           REGION Request selector
               //set Index and RecordLen based on the request
               IF #statParameterPage0 THEN
                   #statIndex := #INDEX_DIRECT_PARAM0;
                   #statRecordLen := #LENGTH_DIRECT_PARAM0;
               ELSIF #statSystemCommands THEN
                   #statIndex := #INDEX_SYSTEM_COMMANDS;
                   #statRecordLen := #LENGTH_SYSTEM_COMMANDS;
               ELSIF #statVendorName THEN
                   #statIndex := #INDEX_VENDOR_NAME;
                   #statRecordLen := #LENGTH_VENDOR_NAME;
               ELSIF #statVendorText THEN
                   #statIndex := #INDEX_VENDOR_TEXT;
                   #statRecordLen := #LENGTH_VENDOR_TEXT;
               ELSIF #statProductName THEN
                   #statIndex := #INDEX_PRODUCT_NAME;
                   #statRecordLen := #LENGTH_PRODUCT_NAME;
               ELSIF #statProductID THEN
                   #statIndex := #INDEX_PRODUCT_ID;
                   #statRecordLen := #LENGTH_PRODUCT_ID;
               ELSIF #statHwRevision THEN
                   #statIndex := #INDEX_HARDWARE_REVISION;
                   #statRecordLen := #LENGTH_HARDWARE_REVISION;
               ELSIF #statFwRevision THEN
                   #statIndex := #INDEX_FIRMWARE_REVISION;
                   #statRecordLen := #LENGTH_FIRMWARE_REVISION;
               ELSIF #statAppSpecificName THEN
                   #statIndex := #INDEX_APP_SPECIFIC_NAME;
                   #statRecordLen := #LENGTH_APP_SPECIFIC_NAME;
               ELSIF #statDiagnosis THEN
                   #statIndex := #INDEX_DIAGNOSTICS;
                   #statRecordLen := #LENGTH_DIAGNOSTICS;
               ELSIF #statMeasurements THEN
                   #statIndex := #INDEX_MEASUREMENTS;
                   #statRecordLen := #LENGTH_MEASUREMENTS;
               ELSIF #statParameters THEN
                   #statIndex := #INDEX_PARAMETERS;
                   #statRecordLen := #LENGTH_PARAMETERS;
               ELSE
                   RETURN;
               END_IF;
           END_REGION

           IF #statReadWrite = #MODE_WRITE THEN
               //prepare statRecord in case of a writing request
               REGION write
                   IF #statSystemCommands THEN
                       #statRecord[0] := #data.systemCommands;

                   ELSIF #statAppSpecificName THEN
                       Strg_TO_Chars(Strg := #data.appSpecificName,
                                     pChars := 0,
                                     Cnt => #tempLen,
                                     Chars := #statRecord);

                       // Fill remaining characters with null
                       FOR #tempIndex := UINT_TO_INT(#tempLen) TO #statRecordLen - 1 DO
                           #statRecord[#tempIndex] := CHAR_TO_BYTE(#EMPTY_CHAR);
                       END_FOR;

                   ELSIF #statParameters THEN
                       #tempRetValSerialize := Serialize(SRC_VARIABLE := #data.parameters, DEST_ARRAY => #tempFieldParameters, POS := #tempPosSerialize);
                       UMOVE_BLK(IN := #tempFieldParameters[0],
                                 COUNT := INT_TO_ULINT(#statRecordLen),
                                 OUT => #statRecord[0]);
                   ELSE    // all other data set are read only
                       ;
                   END_IF;
                   #tempInternalError := #tempRetValSerialize <> WORD_TO_INT(#STATUS_EXECUTION_FINISHED);
               END_REGION

           END_IF;
       END_IF;
   END_REGION

   REGION CALL
       //IOL-Call -> Request to read/write from an IO-Link-Device
       #instDevice(execute := #execute,
                   hwID := #statHwID,
                   cap := #statCap,
                   readWrite := #statReadWrite,
                   "port" := #statPort,
                   pollingPeriod := #statPollingPeriod,
                   index := #statIndex,
                   subindex := #statSubindex,
                   writeLen := #statRecordLen,
                   timeout := #DEVICE_TIMEOUT,
                   record := #statRecord);
   END_REGION

   REGION READ
       // Copy data if available and valid
       IF #instDevice.done = TRUE AND #statDoneOld = FALSE AND #statReadWrite = #MODE_READ THEN
           IF #statParameterPage0 THEN
               UMOVE_BLK(IN := #statRecord[0],
                         COUNT := INT_TO_ULINT(#statRecordLen),
                         OUT => #tempFieldParameterPage0[0]);
               #tempRetValDeserialize := Deserialize(SRC_ARRAY := #tempFieldParameterPage0, DEST_VARIABLE => #data.parameterPage0, POS := #tempPosDeserialize);
           ELSIF #statVendorName THEN
               Chars_TO_Strg(Chars := #statRecord,
                             pChars := 0,
                             Cnt := INT_TO_UINT(#statRecordLen),
                             Strg => #data.vendorName);
           ELSIF #statVendorText THEN
               Chars_TO_Strg(Chars := #statRecord,
                             pChars := 0,
                             Cnt := INT_TO_UINT(#statRecordLen),
                             Strg => #data.vendorText);
           ELSIF #statProductName THEN
               Chars_TO_Strg(Chars := #statRecord,
                             pChars := 0,
                             Cnt := INT_TO_UINT(#statRecordLen),
                             Strg => #data.productName);
           ELSIF #statProductID THEN
               Chars_TO_Strg(Chars := #statRecord,
                             pChars := 0,
                             Cnt := INT_TO_UINT(#statRecordLen),
                             Strg => #data.productID);
           ELSIF #statHwRevision THEN
               Chars_TO_Strg(Chars := #statRecord,
                             pChars := 0,
                             Cnt := INT_TO_UINT(#statRecordLen),
                             Strg => #data.hwRevision);
           ELSIF #statFwRevision THEN
               Chars_TO_Strg(Chars := #statRecord,
                             pChars := 0,
                             Cnt := INT_TO_UINT(#statRecordLen),
                             Strg => #data.fwRevision);
           ELSIF #statAppSpecificName THEN
               Chars_TO_Strg(Chars := #statRecord,
                             pChars := 0,
                             Cnt := INT_TO_UINT(#statRecordLen),
                             Strg => #data.appSpecificName);
           ELSIF #statDiagnosis THEN
               UMOVE_BLK(IN := #statRecord[0],
                         COUNT := INT_TO_ULINT(#statRecordLen),
                         OUT => #tempFieldDiagnostics[0]);
               #tempRetValDeserialize := Deserialize(SRC_ARRAY := #tempFieldDiagnostics, DEST_VARIABLE => #data.diagnostics, POS := #tempPosDeserialize);
           ELSIF #statMeasurements THEN
               UMOVE_BLK(IN := #statRecord[0],
                         COUNT := INT_TO_ULINT(#statRecordLen),
                         OUT => #tempFieldMeasurements[0]);
               #tempRetValDeserialize := Deserialize(SRC_ARRAY := #tempFieldMeasurements, DEST_VARIABLE => #data.measuredValues, POS := #tempPosDeserialize);
           ELSIF #statParameters THEN
               UMOVE_BLK(IN := #statRecord[0],
                         COUNT := INT_TO_ULINT(#statRecordLen),
                         OUT => #tempFieldParameters[0]);
               #tempRetValDeserialize := Deserialize(SRC_ARRAY := #tempFieldParameters, DEST_VARIABLE => #data.parameters, POS := #tempPosDeserialize);
           ELSE  // Other data sets are not defined
               ;
           END_IF;
           #tempInternalError := #tempRetValDeserialize <> WORD_TO_INT(#STATUS_EXECUTION_FINISHED);
       END_IF;

       #statDoneOld := #instDevice.done;
   END_REGION

   REGION OUTPUTS
       IF #tempInternalError THEN //Error occured
           #done := false;
           #busy := false;
           #error := true;
           #status := #ERR_INCONSISTENT_DATA;
       ELSE //Execute successful
           #done := #instDevice.done;
           #busy := #instDevice.busy;
           #error := #instDevice.error;
           #status := #instDevice.status;
           #diagnostics := #instDevice.diagnostics;
       END_IF;
   END_REGION
END_FUNCTION_BLOCK

// folder: LIOLink/S7-1200/1500/Device-specific blocks/SIRIUS/SIRIUS WD

FUNCTION_BLOCK "LIOLink_8WD46"   // FB2, SCL
TITLE = LIOLink_8WD46
{ S7_Optimized_Access := 'TRUE' }
FAMILY : LIOLink
VERSION : 1.0
// Capsule block to communicate with 8WD46
   VAR_INPUT
      execute : Bool;   // Request to execute function
      hwID : HW_IO;   // Hardware identifier of IO-Link master module or first sub module
      cap : Int;   // Client Access Point (CAP) 0xB400 or 0x00E3 (227)
      readWrite : Bool;   // FALSE: read, TRUE: write
      port : Int;   // Port of the IO-Link Master for the Device
      pollingPeriod : Time := T#100MS;   // Time period of polling
      systemCommands : Bool;   // Write system commands
      vendorName : Bool;   // Read Vendor Name
      vendorText : Bool;   // Read Vendor Text
      productName : Bool;   // Read Product Name
      productID : Bool;   // Read Product ID
      productText : Bool;   // Read Product Text
      hwRevision : Bool;   // Read Hardware revision
      fwRevision : Bool;   // Read firmware revision
      appSpecificName : Bool;   // Read/Write Application Specific Name
      functionTag : Bool;   // Read/Write: function tag
      locationTag : Bool;   // Read/Write: location tag
      opHour : Bool;   // Read operating hour
      operatingMode : Bool;   // Read/Write: operating mode (signal mode, auto scale mode, ...)
      lightEffect : USInt;   // Read/Write light effect - 1 to 15: select segment
      soundMode : USInt;   // Read ID of the inserted ID key
      powerReduction : Bool;   // Read/Write power reduction (0: on / 1: off)
      fillLevelMode : Bool;   // Read/Write only in level mode (0: use settings of segment 1-9,15 / 1: use settings of segment 1 )
      headlong : Bool;   // Read/Write orientation of installation (normal / overhead)
      elementCount : Bool;   // Read/Write number of elements
   END_VAR
   VAR_OUTPUT
      done : Bool;   // TRUE: Commanded functionality has been completed successfully
      busy : Bool;   // TRUE: FB is not finished and new output values can be expected
      error : Bool;   // TRUE: An error occurred during the execution of the FB
      status : Word;   // 16#0000 - 16#7FFF: Status of the FB, 16#8000 - 16#FFFF: Error identification
      diagnostics : "LIOLink_typeDiagnostics";   // Diagnostics information of LIOLink_Device
   END_VAR
   VAR_IN_OUT
      data : "LIOLink_8WD46_typeAll";   // Data area, device specific (Data Type)
   END_VAR
   VAR
      instDevice : "LIOLink_Device";
      statRecord : Array[0..#UPPER_BOUND_RECORD] of Byte;   // Record buffer
      statIndex : Int;   // Requested index
      statSubindex : Int;   // Requested subindex
      statRecordLen : Int;   // Length of record to be written
      statHwID : HW_IO;   // Static value for input 'hwID'
      statCap : Int;   // Static value for input 'cap'
      statReadWrite : Bool;   // Static value for input 'readWrite'
      statPort : Int;   // Static value for input 'port'
      statPollingPeriod : Time;   // Static value for input 'pollingPeriod'
      statSystemCommands : Bool;   // Static value for input 'systemCommands'
      statVendorName : Bool;   // Static value for input 'vendorName'
      statVendorText : Bool;   // Static value for input 'vendorText'
      statProductName : Bool;   // Static value for input 'productName'
      statProductID : Bool;   // Static value for input 'productID'
      statProductText : Bool;   // Static value for input 'productText'
      statHwRevision : Bool;   // Static value for input 'hwRevision'
      statFwRevision : Bool;   // Static value for input 'fwRevision'
      statAppSpecificName : Bool;   // Static value for input 'appSpecificName'
      statFunctionTag : Bool;   // Static value for input 'functionTag'
      statLocationTag : Bool;   // Static value for input 'locationTag'
      statOpHour : Bool;   // Static value for input 'opHour'
      statOperatingMode : Bool;   // Static value for input 'operatingMode'
      statLightEffect : USInt;   // Static value for input 'lightEffect'
      statSoundMode : USInt;   // Static value for input 'soundMode'
      statPowerReduction : Bool;   // Static value for input 'powerReduction'
      statFillLevelMode : Bool;   // Static value for input 'fillLevelMode'
      statHeadlong : Bool;   // Static value for input 'headLong'
      statElementCount : Bool;   // Static value for input 'elementCount'
      statRequest : Int;   // Case of request (data set)
      statDoneOld : Bool;   // Last cycle's value of instDevice.done
   END_VAR
   VAR_TEMP
      tempIndex : Int;   // Loop index
      tempLen : UInt;   // Length
      tempRetValSerialize : Int;   // Auxiliary tag for Serialize RetVal
      tempRetValDeserialize : Int;   // Auxiliary tag for Deserialize RetVal
      tempPosSerialize : DInt;   // Auxiliary tag for Serialize POS Output
      tempPosDeserialize : DInt;   // Auxiliary tag for Deserialize POS Output
      tempFieldLightEffects : Array[0..#UPPER_BOUND_LIGHT_EFFECTS] of Byte;   // Auxiliary tag for Light Effects record conversion
      tempFieldSoundMode : Array[0..#UPPER_BOUND_SOUND_MODE] of Byte;   // Auxiliary tag for Sound Mode record conversion
      tempFieldOpHour : Array[0..#UPPER_BOUND_OP_HOUR] of Byte;   // Auxiliary tag for Op Hour record conversion
      tempFieldDiagnostics : Array[0..#UPPER_BOUND_DIAGNOSTICS] of Byte;   // Auxiliary tag for Diagnostics record conversion
      tempInternalError : Bool;   // Auxiliary tag to collect serialize and Deserialize issues
   END_VAR
   VAR CONSTANT
      UPPER_BOUND_RECORD : Int := 231;   // Upper Bound of record buffer
      HIGHEST_REQUEST_NUMBER : Int := 28;   // Highest available request number
      UPPER_BOUND_LIGHT_EFFECTS : Int := 7;   // Upper Bound of Light Effects auxiliary field
      UPPER_BOUND_SOUND_MODE : Int := 15;   // Upper Bound of Sound Mode auxiliary field
      UPPER_BOUND_OP_HOUR : Int := 3;   // Upper Bound of Op Hours auxiliary field
      UPPER_BOUND_DIAGNOSTICS : Int := 19;   // Upper Bound of Diagnostics auxiliary field
      MODE_READ : Bool := FALSE;   // Mode to read data
      MODE_WRITE : Bool := TRUE;   // Mode to write data
      STATUS_IDLE : Word := 16#7000;   // Status: Idle
      STATUS_EXECUTION_FINISHED : Word := 16#0000;   // Execution finished without errors
      ERR_INCONSISTENT_DATA : Word := 16#8402;   // Error: Read data record doesn't match request
      INDEX_SYSTEM_COMMANDS : Int := 2;   // Record Index
      INDEX_VENDOR_NAME : Int := 16;   // Record Index
      INDEX_VENDOR_TEXT : Int := 17;   // Record Index
      INDEX_PRODUCT_NAME : Int := 18;   // Record Index
      INDEX_PRODUCT_ID : Int := 19;   // Record Index
      INDEX_PRODUCT_TEXT : Int := 20;   // Record Index
      INDEX_HARDWARE_REVISION : Int := 22;   // Record Index
      INDEX_FIRMWARE_REVISION : Int := 23;   // Record Index
      INDEX_APP_SPECIFIC_NAME : Int := 24;   // Record Index
      INDEX_FUNCTION_TAG : Int := 25;   // Record Index
      INDEX_LOCATION_TAG : Int := 26;   // Record Index
      INDEX_OPERATING_HOURS : Int := 74;   // Record Index
      INDEX_OPERATING_MODE : Int := 100;   // Record Index
      INDEX_LIGHT_EFFECT : Int := 101;   // Record Index - start of range
      SEGMENT_COUNT_MAX : Int := 15;   // maximum count of segments
      INDEX_SOUND_MODE : Int := 120;   // Record Index - start of range
      SOUND_COUNT_MAX : Int := 10;   // maximum count of sound types
      INDEX_POWER_REDUCTION : Int := 131;   // Record Index
      INDEX_FILL_LEVEL_MODE : Int := 132;   // Record Index
      INDEX_HEADLONG : Int := 138;   // Record Index
      INDEX_COUNT_OF_ELEMENTS : Int := 139;   // Record Index
      LENGTH_SYSTEM_COMMANDS : Int := 1;   // Record Length
      LENGTH_VENDOR_NAME : Int := 48;   // Record Length
      LENGTH_VENDOR_TEXT : Int := 48;   // Record Length
      LENGTH_PRODUCT_NAME : Int := 32;   // Record Length
      LENGTH_PRODUCT_ID : Int := 16;   // Record Length
      LENGTH_PRODUCT_TEXT : Int := 64;   // Record Length
      LENGTH_HARDWARE_REVISION : Int := 16;   // Record Length
      LENGTH_FIRMWARE_REVISION : Int := 16;   // Record Length
      LENGTH_APP_SPECIFIC_NAME : Int := 32;   // Record Length
      LENGTH_FUNCTION_TAG : Int := 32;   // Record Length
      LENGTH_LOCATION_TAG : Int := 32;   // Record Length
      LENGTH_OPERATING_HOURS : Int := 4;   // Record Length
      LENGTH_OPERATING_MODE : Int := 1;   // Record Length
      LENGTH_LIGHT_EFFECT : Int := 8;   // Record Length
      LENGTH_SOUND_MODE : Int := 16;   // Record Length
      LENGTH_POWER_REDUCTION : Int := 1;   // Record Length
      LENGTH_FILL_LEVEL_MODE : Int := 1;   // Record Length
      LENGTH_HEADLONG : Int := 1;   // Record Length
      LENGTH_COUNT_OF_ELEMENTS : Int := 1;   // Record Length
      EMPTY_CHAR : Char := '$00';   // Default empty char to fill empty field entries
      DEVICE_TIMEOUT : Time := T#20S;   // Timeout value for the IO-Link Device Instance
   END_VAR
BEGIN
   REGION BLOCK INFO HEADER
       //===============================================================================
       // Siemens / (c)Copyright 2022
       //-------------------------------------------------------------------------------
       // Title:            LIOLink_8WD46
       // Function:         Capsule block to communicate with 8WD46
       // Library:          LIOLink
       // Author:           Siemens Industry Online Support
       // Tested with:      CPU 1513-1 PN FW 2.8
       // Engineering:      TIA Portal V16
       // Restrictions:     --
       // Requirements:     --
       //-------------------------------------------------------------------------------
       // Change log table:
       // Version  | Date       | Expert in charge       | Changes applied
       //----------|------------|------------------------|------------------------------
       // 01.00.00 | 06.10.2022 | SUP SPH                | First release
       //===============================================================================
   END_REGION

   REGION INIT
       IF (#execute = TRUE AND #instDevice.status = #STATUS_IDLE) THEN
           REGION Inputs
               //Save inputs
               #statHwID := #hwID;
               #statCap := #cap;
               #statReadWrite := #readWrite;
               #statPort := #port;
               #statPollingPeriod := #pollingPeriod;
               #statSystemCommands := #systemCommands;
               #statVendorName := #vendorName;
               #statVendorText := #vendorText;
               #statProductName := #productName;
               #statProductID := #productID;
               #statProductText := #productText;
               #statHwRevision := #hwRevision;
               #statFwRevision := #fwRevision;
               #statAppSpecificName := #appSpecificName;
               #statFunctionTag := #functionTag;
               #statLocationTag := #locationTag;
               #statOpHour := #opHour;
               #statOperatingMode := #operatingMode;
               #statLightEffect := #lightEffect;
               #statSoundMode := #soundMode;
               #statPowerReduction := #powerReduction;
               #statFillLevelMode := #fillLevelMode;
               #statHeadlong := #headlong;
               #statElementCount := #elementCount;
           END_REGION

           REGION Request selector
               //set Index and RecordLen based on the request
               IF #statSystemCommands THEN
                   #statIndex := #INDEX_SYSTEM_COMMANDS;
                   #statRecordLen := #LENGTH_SYSTEM_COMMANDS;
               ELSIF #statVendorName THEN
                   #statIndex := #INDEX_VENDOR_NAME;
                   #statRecordLen := #LENGTH_VENDOR_NAME;
               ELSIF #statVendorText THEN
                   #statIndex := #INDEX_VENDOR_TEXT;
                   #statRecordLen := #LENGTH_VENDOR_TEXT;
               ELSIF #statProductName THEN
                   #statIndex := #INDEX_PRODUCT_NAME;
                   #statRecordLen := #LENGTH_PRODUCT_NAME;
               ELSIF #statProductID THEN
                   #statIndex := #INDEX_PRODUCT_ID;
                   #statRecordLen := #LENGTH_PRODUCT_ID;
               ELSIF #statProductText THEN
                   #statIndex := #INDEX_PRODUCT_TEXT;
                   #statRecordLen := #LENGTH_PRODUCT_TEXT;
               ELSIF #statHwRevision THEN
                   #statIndex := #INDEX_HARDWARE_REVISION;
                   #statRecordLen := #LENGTH_HARDWARE_REVISION;
               ELSIF #statFwRevision THEN
                   #statIndex := #INDEX_FIRMWARE_REVISION;
                   #statRecordLen := #LENGTH_FIRMWARE_REVISION;
               ELSIF #statAppSpecificName THEN
                   #statIndex := #INDEX_APP_SPECIFIC_NAME;
                   #statRecordLen := #LENGTH_APP_SPECIFIC_NAME;
               ELSIF #statFunctionTag THEN
                   #statIndex := #INDEX_FUNCTION_TAG;
                   #statRecordLen := #LENGTH_FUNCTION_TAG;
               ELSIF #statLocationTag THEN
                   #statIndex := #INDEX_LOCATION_TAG;
                   #statRecordLen := #LENGTH_LOCATION_TAG;
               ELSIF #statOpHour THEN
                   #statIndex := #INDEX_OPERATING_HOURS;
                   #statRecordLen := #LENGTH_OPERATING_HOURS;
               ELSIF #statOperatingMode THEN
                   #statIndex := #INDEX_OPERATING_MODE;
                   #statRecordLen := #LENGTH_OPERATING_MODE;
               ELSIF #statLightEffect > 0 AND #statLightEffect <= #SEGMENT_COUNT_MAX THEN
                   #statIndex := #INDEX_LIGHT_EFFECT + #statLightEffect - 1;
                   #statRecordLen := #LENGTH_LIGHT_EFFECT;
               ELSIF #statSoundMode > 0 AND #statSoundMode <= #SOUND_COUNT_MAX THEN
                   #statIndex := #INDEX_SOUND_MODE + #statSoundMode - 1;
                   #statRecordLen := #LENGTH_SOUND_MODE;
               ELSIF #statPowerReduction THEN
                   #statIndex := #INDEX_POWER_REDUCTION;
                   #statRecordLen := #LENGTH_POWER_REDUCTION;
               ELSIF #statFillLevelMode THEN
                   #statIndex := #INDEX_FILL_LEVEL_MODE;
                   #statRecordLen := #LENGTH_FILL_LEVEL_MODE;
               ELSIF #statHeadlong THEN
                   #statIndex := #INDEX_HEADLONG;
                   #statRecordLen := #LENGTH_HEADLONG;
               ELSIF #statElementCount THEN
                   #statIndex := #INDEX_COUNT_OF_ELEMENTS;
                   #statRecordLen := #LENGTH_COUNT_OF_ELEMENTS;
               ELSE
                   RETURN;
               END_IF;
           END_REGION

           IF #statReadWrite = #MODE_WRITE THEN
               //prepare statRecord in case of a writing request
               REGION write
                   IF #statSystemCommands THEN
                       #statRecord[0] := #data.systemCommand;

                   ELSIF #statAppSpecificName THEN
                       Strg_TO_Chars(Strg := #data.appSpecificName,
                                     pChars := 0,
                                     Cnt => #tempLen,
                                     Chars := #statRecord);

                       // Fill remaining characters with null
                       FOR #tempIndex := UINT_TO_INT(#tempLen) TO #statRecordLen - 1 DO
                           #statRecord[#tempIndex] := CHAR_TO_BYTE(#EMPTY_CHAR);
                       END_FOR;

                   ELSIF #statFunctionTag THEN
                       Strg_TO_Chars(Strg := #data.functionTag,
                                     pChars := 0,
                                     Cnt => #tempLen,
                                     Chars := #statRecord);

                       // Fill remaining characters with null
                       FOR #tempIndex := UINT_TO_INT(#tempLen) TO #statRecordLen - 1 DO
                           #statRecord[#tempIndex] := CHAR_TO_BYTE(#EMPTY_CHAR);
                       END_FOR;

                   ELSIF #statLocationTag THEN
                       Strg_TO_Chars(Strg := #data.locationTag,
                                     pChars := 0,
                                     Cnt => #tempLen,
                                     Chars := #statRecord);

                       // Fill remaining characters with null
                       FOR #tempIndex := UINT_TO_INT(#tempLen) TO #statRecordLen - 1 DO
                           #statRecord[#tempIndex] := CHAR_TO_BYTE(#EMPTY_CHAR);
                       END_FOR;

                   ELSIF #statOperatingMode THEN
                       #statRecord[0] := #data.operatingMode;

                   ELSIF #statLightEffect > 0 AND #statLightEffect <= #SEGMENT_COUNT_MAX THEN
                       #tempRetValSerialize := Serialize(SRC_VARIABLE := #data.lightEffects[#statLightEffect], DEST_ARRAY => #tempFieldLightEffects, POS := #tempPosSerialize);
                       UMOVE_BLK(IN := #tempFieldLightEffects[0],
                                 COUNT := INT_TO_ULINT(#statRecordLen),
                                 OUT => #statRecord[0]);

                   ELSIF #statSoundMode > 0 AND #statSoundMode <= #SOUND_COUNT_MAX THEN
                       #statRecord[0] := #data.soundMode[#statSoundMode].mode;
                       #statRecord[1] := #data.soundMode[#statSoundMode].frequency1Start.%B1;
                       #statRecord[2] := #data.soundMode[#statSoundMode].frequency1Start.%B0;
                       #statRecord[3] := #data.soundMode[#statSoundMode].frequency2Stop.%B1;
                       #statRecord[4] := #data.soundMode[#statSoundMode].frequency2Stop.%B0;
                       #statRecord[5] := #data.soundMode[#statSoundMode].frequency1Periode.%B1;
                       #statRecord[6] := #data.soundMode[#statSoundMode].frequency1Periode.%B0;
                       #statRecord[7] := #data.soundMode[#statSoundMode].volume;
                       #statRecord[8] := #data.soundMode[#statSoundMode].count.%B1;
                       #statRecord[9] := #data.soundMode[#statSoundMode].count.%B0;
                       #statRecord[10] := #data.soundMode[#statSoundMode].brakeToRepeat.%B1;
                       #statRecord[11] := #data.soundMode[#statSoundMode].brakeToRepeat.%B0;
                       #statRecord[12] := #data.soundMode[#statSoundMode].BrakeBetweenCycles.%B1;
                       #statRecord[13] := #data.soundMode[#statSoundMode].BrakeBetweenCycles.%B0;
                       #statRecord[14] := #data.soundMode[#statSoundMode].holdingPeriodeFrequency2.%B1;
                       #statRecord[15] := #data.soundMode[#statSoundMode].holdingPeriodeFrequency2.%B0;

                   ELSIF #statPowerReduction THEN
                       #statRecord[0] := #data.#powerReduction;

                   ELSIF #statFillLevelMode THEN
                       #statRecord[0] := #data.fillLevelMode;

                   ELSIF #statHeadlong THEN
                       #statRecord[0] := #data.headlong;

                   ELSIF #statElementCount THEN
                       #statRecord[0] := #data.elementCount;

                   ELSE // All other data sets are read only  
                       ;
                   END_IF;
                   #tempInternalError := #tempRetValSerialize <> WORD_TO_INT(#STATUS_EXECUTION_FINISHED);
               END_REGION
           END_IF;
       END_IF;
   END_REGION

   REGION CALL
       //IOL-Call -> Request to read/write from an IO-Link-Device
       #instDevice(execute := #execute,
                   hwID := #statHwID,
                   cap := #statCap,
                   readWrite := #statReadWrite,
                   "port" := #statPort,
                   pollingPeriod := #statPollingPeriod,
                   index := #statIndex,
                   subindex := #statSubindex,
                   writeLen := #statRecordLen,
                   timeout := #DEVICE_TIMEOUT,
                   record := #statRecord);
   END_REGION

   REGION READ
       // Copy data if available and valid
       IF #instDevice.done = TRUE AND #statDoneOld = FALSE AND #statReadWrite = #MODE_READ THEN
           IF #statVendorName THEN
               Chars_TO_Strg(Chars := #statRecord,
                             pChars := 0,
                             Cnt := INT_TO_UINT(#statRecordLen),
                             Strg => #data.vendorName);

           ELSIF #statVendorText THEN
               Chars_TO_Strg(Chars := #statRecord,
                             pChars := 0,
                             Cnt := INT_TO_UINT(#statRecordLen),
                             Strg => #data.vendorText);

           ELSIF #statProductName THEN
               Chars_TO_Strg(Chars := #statRecord,
                             pChars := 0,
                             Cnt := INT_TO_UINT(#statRecordLen),
                             Strg => #data.productName);

           ELSIF #statProductID THEN
               Chars_TO_Strg(Chars := #statRecord,
                             pChars := 0,
                             Cnt := INT_TO_UINT(#statRecordLen),
                             Strg => #data.productId);

           ELSIF #statProductText THEN
               Chars_TO_Strg(Chars := #statRecord,
                             pChars := 0,
                             Cnt := INT_TO_UINT(#statRecordLen),
                             Strg => #data.productText);

           ELSIF #statHwRevision THEN
               Chars_TO_Strg(Chars := #statRecord,
                             pChars := 0,
                             Cnt := INT_TO_UINT(#statRecordLen),
                             Strg => #data.hwRevision);

           ELSIF #statFwRevision THEN
               Chars_TO_Strg(Chars := #statRecord,
                             pChars := 0,
                             Cnt := INT_TO_UINT(#statRecordLen),
                             Strg => #data.fwRevision);

           ELSIF #statAppSpecificName THEN
               Chars_TO_Strg(Chars := #statRecord,
                             pChars := 0,
                             Cnt := INT_TO_UINT(#statRecordLen),
                             Strg => #data.appSpecificName);

           ELSIF #statFunctionTag THEN
               Chars_TO_Strg(Chars := #statRecord,
                             pChars := 0,
                             Cnt := INT_TO_UINT(#statRecordLen),
                             Strg => #data.#functionTag);

           ELSIF #statLocationTag THEN
               Chars_TO_Strg(Chars := #statRecord,
                             pChars := 0,
                             Cnt := INT_TO_UINT(#statRecordLen),
                             Strg => #data.#locationTag);

           ELSIF #statOpHour THEN
               UMOVE_BLK(IN := #statRecord[0],
                         COUNT := INT_TO_ULINT(#statRecordLen),
                         OUT => #tempFieldOpHour[0]);
               #tempRetValDeserialize := Deserialize(SRC_ARRAY := #tempFieldOpHour, DEST_VARIABLE => #data.opHour, POS := #tempPosDeserialize);

           ELSIF #statLightEffect > 0 AND #statLightEffect <= #SEGMENT_COUNT_MAX THEN
               UMOVE_BLK(IN := #statRecord[0],
                         COUNT := INT_TO_ULINT(#statRecordLen),
                         OUT => #tempFieldLightEffects[0]);
               #tempRetValDeserialize := Deserialize(SRC_ARRAY := #tempFieldLightEffects, DEST_VARIABLE => #data.lightEffects[#statLightEffect], POS := #tempPosDeserialize);

           ELSIF #statSoundMode > 0 AND #statSoundMode <= #SOUND_COUNT_MAX THEN
               #data.soundMode[#statSoundMode].mode := #statRecord[0];
               #data.soundMode[#statSoundMode].frequency1Start.%B0 := #statRecord[2];
               #data.soundMode[#statSoundMode].frequency1Start.%B1 := #statRecord[1];
               #data.soundMode[#statSoundMode].frequency2Stop.%B0 := #statRecord[4];
               #data.soundMode[#statSoundMode].frequency2Stop.%B1 := #statRecord[3];
               #data.soundMode[#statSoundMode].frequency1Periode.%B0 := #statRecord[6];
               #data.soundMode[#statSoundMode].frequency1Periode.%B1 := #statRecord[5];
               #data.soundMode[#statSoundMode].volume := #statRecord[7];
               #data.soundMode[#statSoundMode].count.%B0 := #statRecord[9];
               #data.soundMode[#statSoundMode].count.%B1 := #statRecord[8];
               #data.soundMode[#statSoundMode].brakeToRepeat.%B0 := #statRecord[11];
               #data.soundMode[#statSoundMode].brakeToRepeat.%B1 := #statRecord[10];
               #data.soundMode[#statSoundMode].BrakeBetweenCycles.%B0 := #statRecord[13];
               #data.soundMode[#statSoundMode].BrakeBetweenCycles.%B1 := #statRecord[12];
               #data.soundMode[#statSoundMode].holdingPeriodeFrequency2.%B0 := #statRecord[15];
               #data.soundMode[#statSoundMode].holdingPeriodeFrequency2.%B1 := #statRecord[14];


           ELSIF #statPowerReduction THEN
               #data.powerReduction := #statRecord[0];

           ELSIF #statFillLevelMode THEN
               #data.#fillLevelMode := #statRecord[0];

           ELSIF #statHeadlong THEN
               #data.#headlong := #statRecord[0];

           ELSIF #statElementCount THEN
               #data.elementCount := #statRecord[0];
           ELSE // Other data sets are not defined
               ;
           END_IF;
           #tempInternalError := #tempRetValDeserialize <> WORD_TO_INT(#STATUS_EXECUTION_FINISHED);
       END_IF;

       #statDoneOld := #instDevice.done;
   END_REGION

   REGION OUTPUTS
       IF #tempInternalError THEN //Error occured
           #done := false;
           #busy := false;
           #error := true;
           #status := #ERR_INCONSISTENT_DATA;
       ELSE //Execute successful
           #done := #instDevice.done;
           #busy := #instDevice.busy;
           #error := #instDevice.error;
           #status := #instDevice.status;
           #diagnostics := #instDevice.diagnostics;
       END_IF;
   END_REGION
END_FUNCTION_BLOCK

// folder: LIOLink/S7-1200/1500/Profile blocks

FUNCTION_BLOCK "LIOLink_MultiAdjSwitchingSensor"   // FB8, SCL
TITLE = LIOLink_MultiAdjSwitchingSensor
{ S7_Optimized_Access := 'TRUE' }
AUTHOR : SUP_Applications
FAMILY : LIOLink
VERSION : 2.0
// Provides a standardized interface and access method for parameterization of a sensor using the Smart Sensor profile. In particular, the FB can be used by sensors that can be assigned to the measuring device profile type 2, i.e. IO Link Devices that support the smart sensor profile "Multiple Adjustable Switching Sensors".
   VAR_INPUT
      execute : Bool;   // Execute selected function
      hwID : HW_IO;   // Hardware identifier of IO-Link master module (sub module for ET 200eco PN)
      cap : Int;   // Client Access Point; 0xB400 for ET 200eco PN, CM 8x IO-Link, else 0xE003 (227)
      port : Int;   // Port on IO-Link master module
      backupEnable : Bool;   // TRUE: Data storage enabled, FALSE: disabled
      function : Int;   // 0: no_func, 1: rd_all, 2: wr_conf, 3: wr_param, 4: teach
      logicIn : Bool;   // This variable defines the value for a new Switchpoint to be written to the sensor on a Request with Function ‘wr_conf’
      setpointIn1 : Int;   // This variable defines the value for a new Setpoint to be written to the sensor on a Request with Function ‘wr_param’
      setpointIn2 : Int;   // This variable defines the value for a new Setpoint to be written to the sensor on a Request with Function ‘wr_param’
      teachMode : Int;   // 0: no_teach, 1: single_value, 2: two_value, 3: dynamic
      teachTimer : Time;   // Defines the duration of the dynamic teach time
      applyAuto : Bool;   // Teaching result is applied automatically after two teach points were teached (only applies to two value teach mode)
      teachRequest : Bool;   // A rising edge triggers one step of teach process to be executed according to the selected function at input teachFunction
      teachFunction : Int;   // 0: no teach, 1: teach 1; 2: teach 2; 3: apply; 4: abort
   END_VAR
   VAR_OUTPUT
      done : Bool;   // The signal is set, if the FB has completed a requested operation.
      busy : Bool;   // The signal is set, if the FB is executing a requested operation.
      error : Bool;   // The signal is set, if an error occurred during execution of a requested operation.
      status : Word := 16#7000;   // Provides block internal status
      diagnostics : "LIOLink_typeDiagnostics";   // Diagnostics information of LIOLink_Device
      logicOut : Bool;   // Represents the current value of the parameter Logic from the sensor.
      setpointOut1 : Int;   // represents the current value of the parameter Setpoint from the sensor.
      setpointOut2 : Int;   // represents the current value of the parameter Setpoint from the sensor.
      permitTeach1 : Bool;   // The signal is set, if a teach request for teach function ‘teach_1’ is allowed
      permitTeach2 : Bool;   // The signal is set, if a teach request for teach function ‘teach_2’ is allowed
      permitApply : Bool;   // The signal is set, if a teach request for teach function ‘apply’ is allowed
      permitAbort : Bool;   // The signal is set, if a teach request for teach function ‘abort’ is allowed
   END_VAR
   VAR
      statExecuteOld : Bool;   // Old value of 'execute' input for edge detection
      statDone : Bool;   // Static value for output 'done'
      statBusy : Bool;   // Static value for output 'busy'
      statError : Bool;   // Static value for output 'error'
      statStatus : Word := 16#7000;   // Static value for output 'status'
      statSubfunctionStatus : Word;   // Status or return value of called FBs, FCs and system blocks
      statFBState : Int;   // State of the state machine
      statFBSubState : Int;   // Sub state of the state machine
      statFBErrorState : DInt;   // State in the state machine of the block where the error occurred
      statEmptyDiagnostics : "LIOLink_typeDiagnostics";   // Empty diagnostics information (for initialization purposes only)
      statTeachRequestOld : Bool;   // Used to check TeachRequest Input for rising edge
      statRwRecordIOLData : Array[0..231] of Byte;   // Buffer, used to work with IO_Link_Device
      instDevice : "LIOLink_Device";
      statIndexRead : Int;   // Used to address the index which has to be read next
      statLenRead : Int;   // Used to handle the length of the parameter which has to be read next
      statTP1Teached : Bool;   // Is set after tp1 of two value teach has been teached
      statTP2Teached : Bool;   // Is set after tp2 of two value teach has been teached
      instTimer : TON_TIME;   // Timer for dynamic teach
      statTeachStarted : Bool;   // Help variable to determine if dynamic each has been started
      statMyPermitTeach1 : Bool;   // Help variable for internal handling of PermitTeach1
      statMyPermitTeach2 : Bool;   // Help variable for internal handling of PermitTeach2
      statMyPermitApply : Bool;   // Help variable for internal handling of PermitTeachApply
      statMyPermitAbort : Bool;   // Help variable for internal handling of PermitTeachAbort
   END_VAR
   VAR_TEMP
      tempExecute : Bool;   // Temporary value for input 'execute'
      tempSetpointOut1 : Word;   // Temporary variable to encode the output "setpointOut" in byte
      tempSetpointIn1 : Word;   // Temporary variable to encode the Input "setpointIn" in byte
      tempSetpointOut2 : Word;   // Temporary variable to encode the output "setpointOut" in byte
      tempSetpointIn2 : Word;   // Temporary variable to encode the Input "setpointIn" in byte
   END_VAR
   VAR CONSTANT
      MODE_READ : Bool;   // Mode to read data
      MODE_WRITE : Bool := TRUE;   // Mode to write data
      FB_STATE_NO_PROCESSING : Int;   // Idle State
      FB_STATE_READ_ALL : Int := 102;   // State to read Setpoint and SwitchPointLogic
      FB_STATE_WRITE_CONF : Int := 103;   // State to write SwitchPointLogic
      FB_STATE_WRITE_PARAM : Int := 104;   // State to write Setpoint
      FB_STATE_BACKUP : Int := 105;   // State to trigger Datastorage mechanism
      FB_STATE_CHECK_TEACH_STATE : Int := 201;   // State to check current teach state before starting teach-in process
      FB_STATE_CHECK_TEACH_MODE : Int := 202;   // State to determine which teach mode is intended (sigle value, two value, dynamic)
      FB_STATE_SINGLE_VAL_TEACH_IN : Int := 210;   // State for teaching single value teach
      FB_STATE_TWO_VAL_TEACH_IN : Int := 220;   // State for teaching two value teach
      FB_SUB_STATE_TWO_VAL_UPDATE_STATUS : Int := 221;   // Sub state inside two value teach to check TI_Result during two value teach
      FB_SUB_STATE_TWO_VAL_WRITE_COMMAND : Int := 222;   // Sub state inside two value teach to write teach commands during two value teach
      FB_STATE_DYNAMIC_TEACH_IN : Int := 230;   // State for teaching dynamic teach
      FB_SUB_STATE_DYNAMIC_UPDATE_STATUS : Int := 231;   // Sub state inside dynamic teach to check TI_Result during dynamic teach
      FB_SUB_STATE_DYNAMIC_WRITE_COMMAND : Int := 232;   // Sub state inside dynamic teach to write teach commands during dynamic teach
      FB_STATE_CHECK_RESULT : Int := 240;   // State to check result of executed teach mode
      FB_STATE_ABORT_TEACH : Int := 260;   // State to abort teach procedure
      INDEX_SYS_CMD : Int := 2;   // Index of "System command"
      INDEX_SSC_PARAM : Int := 56;   // Index of "SSC Param"
      INDEX_SSC_CONFIG : Int := 57;   // Index of "SSC Config"
      INDEX_TI_RESULT : Int := 59;   // Index of "Teach-in Result"
      TICMD_APPLY : Byte := 16#40;   // Teach-in command "Teach Apply"
      TICMD_TEACH_SP : Byte := 16#41;   // Teach-in command "Teach SP"
      TICMD_TEACH_SP_TP1 : Byte := 16#43;   // Teach-in command "Teach SP TP1"
      TICMD_TEACH_SP_TP2 : Byte := 16#44;   // Teach-in command "Teach SP TP2"
      TICMD_TEACH_SP_START : Byte := 16#47;   // Teach-in command "Teach SP Start"
      TICMD_TEACH_SP_STOP : Byte := 16#48;   // Teach-in command "Teach SP Stop"
      TICMD_TEACH_CANCEL : Byte := 16#4F;   // Teach-in command "Teach cancel"
      MASK_FLAG_TP1 : Byte := 16#10;   // Mask flag SP TP1/Teachpoint successfully acquired
      MASK_FLAG_TP2 : Byte := 16#20;   // Mask flag SP TP2/Teachpoint successfully acquired
      MASK_TEACH_STATE : Byte := 16#0F;   // Mask teach state
      TEACH_STATE_IDLE : Int := 0;   // Constatnt for TI_Result = Idle
      TEACH_STATE_SUCCESS : Int := 1;   // Constatnt for TI_Result = Success
      TEACH_STATE_WAIT_FOR_COMMAND : Int := 4;   // Constatnt for TI_Result = Wait for Command
      TEACH_STATE_BUSY : Int := 5;   // Constatnt for TI_Result = Busy
      TEACH_STATE_ERROR : Int := 7;   // Constatnt for TI_Result = Error
      STATUS_EXECUTION_FINISHED : Word := 16#0000;   // Status: Teach process successfull/ Ready to Start Teach-In process / idle
      STATUS_NO_CALL : Word := 16#7000;   // Status: Function block is idle
      STATUS_BUSY_READING : Word := 16#7011;   // Status: Busy reading data
      STATUS_BUSY_WRITING : Word := 16#7012;   // Status: Busy writing data
      STATUS_BUSY_BACKUP : Word := 16#7026;   // Status: Busy with backup
      STATUS_TEACH_STARTED : Word := 16#7101;   // Status: Teach-in process started
      STATUS_TEACH_SUBSEQUENT_CALL : Word := 16#7102;   // Status: Teach-in process subsequent call
      STATUS_TEACH_SINGLE_WAITING : Word := 16#7110;   // Status: Teach-in process for single value teach-in is waiting for further command
      STATUS_TEACH_SINGLE_BUSY : Word := 16#7111;   // Status: Teach-in process for single value teach-in is executed
      STATUS_TEACH_TWO_WAITING : Word := 16#7120;   // Status: Two value teach-in process is waiting for further command
      STATUS_TEACH_TWO_BUSY : Word := 16#7121;   // Status: Two value teach-in process is being executed
      STATUS_TEACH_DYNAMIC_WAITING : Word := 16#7130;   // Status: Dynamic teach-in process is waiting for further command
      STATUS_TEACH_DYNAMIC_BUSY : Word := 16#7131;   // Status: Dynamic teach-in process is being executed
      STATUS_TEACH_WAITING_APPLY : Word := 16#7140;   // Status: Teach-in process is waiting for apply action command
      STATUS_TEACH_APPLYING : Word := 16#7141;   // Status: Teach-in process is executed, perform action
      STATUS_TEACH_ABORTING : Word := 16#7151;   // Status: Teach-in process is executed, abort action
      SUB_STATUS_NO_ERROR : Word := 16#0000;   // No error occured in subfunction call
      ERR_UNKNOWN_FUNCTION : Word := 16#8030;   // Error: Selected function unknown
      ERR_TEACH_DEVICE : Word := 16#8330;   // Error: Device detected an error during the teach-in process
      ERR_TEACH_NOT_ALLOWED : Word := 16#8331;   // Error: Teach function not permitted in this state
      ERR_TEACH_MODE_UNKNOWN : Word := 16#8332;   // Error: Selected teach mode unknown
      ERR_DEVICE_FB : Word := 16#8600;   // Error in LIOLink_Device, see "diagnostics"
      FUNC_NOTHING : Int := 0;   // Execute no function
      FUNC_RD_ALL : Int := 1;   // Function to read logic and setpoint from sensor
      FUNC_WR_CONF : Int := 2;   // Function write logic to sensor
      FUNC_WR_PARAM : Int := 3;   // Function to write setpoint to sensor
      FUNC_TEACH : Int := 4;   // Function to enter the teach operation
      TEACH_MODE_NO_TEACH : Int := 0;   // No teach mode
      TEACH_MODE_SINGLE_VALUE_TEACH_IN : Int := 1;   // Teach Mode Single value teach-in
      TEACH_MODE_TWO_VALUE_TEACH_IN : Int := 2;   // Teach Mode Two value teach-in
      TEACH_MODE_DYNAMIC_TEACH_IN : Int := 3;   // Teach Mode dynamic teach-in
      TEACH_FUNCTION_1 : Int := 1;   // Teach function 1: Start Teach Step 1
      TEACH_FUNCTION_2 : Int := 2;   // Teach function 2: Start Teach Step 2
      TEACH_FUNCTION_APPLY : Int := 3;   // Apply two value teach results
      TEACH_FUNCTION_ABORT : Int := 4;   // Abort of the current teach sequence
   END_VAR
BEGIN
   REGION BLOCK INFO HEADER
       //===============================================================================
       // Siemens / (c)Copyright 2023
       //-------------------------------------------------------------------------------
       // Title:            LIOLink_MultiAdjSwitchingSensor
       // Function:         This FB provides a standardized interface and access method for
       //                   parameterization of a sensor using the Smart Sensor profile.
       //                   In particular, the FB can be used by sensors that can be assigned
       //                   to the measuring device profile type 2, i.e. IO Link Devices that
       //                   support the smart sensor profile "Multiple Adjustable Switching Sensors".
       // Library:          LIOLink
       // Author:           SUP Applications
       // Tested with:      CPU 1513-1 PN FW 2.8
       // Engineering:      TIA Portal V16
       // Restrictions:     --
       // Requirements:     --
       //-------------------------------------------------------------------------------
       // Change log table:
       // Version  | Date       | Expert in charge       | Changes applied
       //----------|------------|------------------------|------------------------------
       // 01.00.00 | 28.02.2023 | SUP Applications       | First release
       //===============================================================================
   END_REGION

   #tempExecute := #execute; // Work with temporary value / create process image

   REGION TRIGGERING
       IF (#tempExecute = TRUE) AND (#statExecuteOld = FALSE) // Check if FB is triggered
           AND (#statStatus = #STATUS_NO_CALL)
       THEN // First call; initialize FB
           #statDone := FALSE;
           #statBusy := TRUE;
           #statError := FALSE;
           #statSubfunctionStatus := #SUB_STATUS_NO_ERROR;
           #statFBErrorState := 0;
           #diagnostics := #statEmptyDiagnostics;

           #statMyPermitAbort := FALSE;
           #statMyPermitApply := FALSE;
           #statMyPermitTeach1 := FALSE;
           #statMyPermitTeach2 := FALSE;


           // Set up LIOLink_Device
           #instDevice(execute := FALSE,
                       hwID := #hwID,
                       cap := #cap,
                       readWrite := 0,
                       "port" := #port,
                       index := 0,
                       subindex := 0,
                       record := #statRwRecordIOLData);

           CASE #function OF
               #FUNC_NOTHING:
                   #statStatus := #STATUS_EXECUTION_FINISHED;

               #FUNC_RD_ALL:
                   #statStatus := #STATUS_BUSY_READING;
                   #statFBState := #FB_STATE_READ_ALL;
                   #statIndexRead := #INDEX_SSC_PARAM;
                   #statLenRead := 2;

               #FUNC_WR_CONF:
                   #statStatus := #STATUS_BUSY_WRITING;
                   #statFBState := #FB_STATE_WRITE_CONF;

               #FUNC_WR_PARAM:
                   #statStatus := #STATUS_BUSY_WRITING;
                   #statFBState := #FB_STATE_WRITE_PARAM;

               #FUNC_TEACH:
                   #statStatus := #STATUS_TEACH_STARTED;
                   #statFBState := #FB_STATE_CHECK_TEACH_STATE;

               ELSE: // Error: not defined
                   #statStatus := #ERR_UNKNOWN_FUNCTION;
           END_CASE;

       ELSIF (#statStatus = #STATUS_TEACH_STARTED) THEN
           #statStatus := #STATUS_TEACH_SUBSEQUENT_CALL;
       END_IF;

       // Edge detection 'execute' input
       #statExecuteOld := #tempExecute;
   END_REGION TRIGGERING

   IF (#statStatus = #STATUS_NO_CALL) THEN // Nothing to do -> End here to reduce "system load"
       RETURN;
   END_IF;

   REGION STATE_MACHINE
       CASE #statFBState OF // State machine of FB
           #FB_STATE_NO_PROCESSING:
               REGION no processing
                   // No processing active
                   ;
               END_REGION no processing

           #FB_STATE_CHECK_TEACH_STATE..#FB_STATE_ABORT_TEACH:
               REGION teach
                   REGION check teach state
                       IF #statFBState = #FB_STATE_CHECK_TEACH_STATE THEN //check Teach status 
                           #instDevice(execute := TRUE,
                                       readWrite := #MODE_READ,
                                       index := #INDEX_TI_RESULT,
                                       record := #statRwRecordIOLData);

                           IF #instDevice.done THEN
                               #instDevice(execute := FALSE,
                                           record := #statRwRecordIOLData);

                               IF (#statRwRecordIOLData[0] AND #MASK_TEACH_STATE) = INT_TO_BYTE(#TEACH_STATE_BUSY) THEN
                                   ; // Keep trying until teach state of device is not busy
                               ELSE
                                   CASE #teachMode OF
                                       #TEACH_MODE_NO_TEACH:
                                           #statStatus := #STATUS_EXECUTION_FINISHED;

                                       #TEACH_MODE_SINGLE_VALUE_TEACH_IN:
                                           #statStatus := #STATUS_TEACH_SINGLE_WAITING;
                                           #statMyPermitTeach1 := TRUE;
                                           #statFBState := #FB_STATE_SINGLE_VAL_TEACH_IN;

                                       #TEACH_MODE_TWO_VALUE_TEACH_IN:
                                           #statStatus := #STATUS_TEACH_TWO_WAITING;
                                           #statTP1Teached := FALSE;
                                           #statTP2Teached := FALSE;
                                           #statMyPermitTeach1 := TRUE;
                                           #statMyPermitTeach2 := TRUE;
                                           #statFBState := #FB_STATE_TWO_VAL_TEACH_IN;
                                           #statFBSubState := 0;

                                       #TEACH_MODE_DYNAMIC_TEACH_IN:
                                           #statStatus := #STATUS_TEACH_DYNAMIC_WAITING;
                                           #statMyPermitTeach1 := TRUE;
                                           #statTeachStarted := FALSE;
                                           #instTimer(PT := #teachTimer,
                                                      IN := FALSE);
                                           #statFBState := #FB_STATE_DYNAMIC_TEACH_IN;
                                           #statFBSubState := 0;

                                       ELSE  // Error: NOT defined
                                           #statStatus := #ERR_TEACH_MODE_UNKNOWN;
                                   END_CASE;
                               END_IF;
                           END_IF;
                       END_IF;
                   END_REGION check teach state

                   REGION single teach-in
                       IF #statFBState = #FB_STATE_SINGLE_VAL_TEACH_IN THEN

                           // Teach SP
                           #statRwRecordIOLData[0] := #TICMD_TEACH_SP;
                           #instDevice(execute := #teachRequest AND NOT #statTeachRequestOld AND #teachFunction = #TEACH_FUNCTION_1,
                                       readWrite := #MODE_WRITE,
                                       index := #INDEX_SYS_CMD,
                                       writeLen := 1,
                                       record := #statRwRecordIOLData);

                           IF #instDevice.busy THEN
                               #statStatus := #STATUS_TEACH_SINGLE_BUSY;
                           ELSIF #instDevice.done THEN
                               #instDevice(execute := FALSE,
                                           record := #statRwRecordIOLData);
                               #statFBState := #FB_STATE_CHECK_RESULT;
                           END_IF;
                       END_IF;
                   END_REGION single teach-in

                   REGION two value teach-in
                       IF #statFBState = #FB_STATE_TWO_VAL_TEACH_IN THEN

                           // Wait for rising edge of teachRequest
                           IF #teachRequest AND NOT #statTeachRequestOld THEN
                               #statStatus := #STATUS_TEACH_TWO_BUSY;

                               IF #teachFunction = #TEACH_FUNCTION_1 THEN
                                   // Teach Point 1
                                   #statRwRecordIOLData[0] := #TICMD_TEACH_SP_TP1;
                               ELSIF #teachFunction = #TEACH_FUNCTION_2 THEN
                                   // Teach Point 2
                                   #statRwRecordIOLData[0] := #TICMD_TEACH_SP_TP2;
                               ELSIF #teachFunction = #TEACH_FUNCTION_APPLY THEN
                                   // Teach Apply
                                   #statRwRecordIOLData[0] := #TICMD_APPLY;
                               END_IF;
                               #statFBSubState := #FB_SUB_STATE_TWO_VAL_WRITE_COMMAND;
                           END_IF;

                           IF #statFBSubState = #FB_SUB_STATE_TWO_VAL_UPDATE_STATUS THEN
                               #instDevice(execute := TRUE,
                                           readWrite := #MODE_READ,
                                           index := #INDEX_TI_RESULT,
                                           record := #statRwRecordIOLData);

                               IF #instDevice.done THEN
                                   #instDevice(execute := FALSE,
                                               record := #statRwRecordIOLData);

                                   // Evaluate response from device
                                   IF (#statRwRecordIOLData[0] AND #MASK_TEACH_STATE) = INT_TO_BYTE(#TEACH_STATE_IDLE) OR
                                       (#statRwRecordIOLData[0] AND #MASK_TEACH_STATE) = INT_TO_BYTE(#TEACH_STATE_SUCCESS)
                                   THEN
                                       #statStatus := #STATUS_TEACH_TWO_BUSY;
                                       #statFBSubState := 0;
                                   ELSIF (#statRwRecordIOLData[0] AND #MASK_TEACH_STATE) = INT_TO_BYTE(#TEACH_STATE_WAIT_FOR_COMMAND) THEN
                                       #statStatus := #STATUS_TEACH_TWO_WAITING;
                                       #statFBSubState := 0;
                                   ELSIF (#statRwRecordIOLData[0] AND #MASK_TEACH_STATE) = INT_TO_BYTE(#TEACH_STATE_BUSY) THEN
                                       #statStatus := #STATUS_TEACH_TWO_BUSY;
                                   ELSIF (#statRwRecordIOLData[0] AND #MASK_TEACH_STATE) = INT_TO_BYTE(#TEACH_STATE_ERROR) THEN
                                       #statStatus := #ERR_TEACH_DEVICE;
                                   END_IF;

                                   // Check if Teachpoints were successfuly acquired
                                   IF (#statRwRecordIOLData[0] AND #MASK_FLAG_TP1) = #MASK_FLAG_TP1 THEN
                                       #statTP1Teached := TRUE;
                                   END_IF;

                                   IF (#statRwRecordIOLData[0] AND #MASK_FLAG_TP2) = #MASK_FLAG_TP2 THEN
                                       #statTP2Teached := TRUE;
                                   END_IF;
                               END_IF;
                           END_IF;

                           // Write Teach Commands
                           IF #statFBSubState = #FB_SUB_STATE_TWO_VAL_WRITE_COMMAND THEN
                               #instDevice(execute := TRUE,
                                           readWrite := #MODE_WRITE,
                                           index := #INDEX_SYS_CMD,
                                           writeLen := 1,
                                           record := #statRwRecordIOLData);

                               IF #instDevice.done THEN
                                   #instDevice(execute := FALSE,
                                               record := #statRwRecordIOLData);
                                   #statFBSubState := #FB_SUB_STATE_TWO_VAL_UPDATE_STATUS;
                                   #statMyPermitAbort := TRUE;

                                   IF #statRwRecordIOLData[0] = #TICMD_APPLY THEN
                                       #statFBState := #FB_STATE_CHECK_RESULT;
                                       #statStatus := #STATUS_TEACH_APPLYING; // Busy, Teach process, apply action
                                   END_IF;
                               END_IF;
                           END_IF;

                           IF #statTP1Teached AND #statTP2Teached THEN
                               #statMyPermitApply := TRUE;

                               IF #applyAuto THEN
                                   #statRwRecordIOLData[0] := #TICMD_APPLY;
                                   #statFBSubState := #FB_SUB_STATE_TWO_VAL_WRITE_COMMAND;
                               END_IF;
                           END_IF;
                       END_IF;
                   END_REGION

                   REGION dynamic teach-in
                       IF #statFBState = #FB_STATE_DYNAMIC_TEACH_IN THEN

                           //Wait for rising edge of TeachRequest input
                           IF #teachRequest AND NOT #statTeachRequestOld THEN
                               #statStatus := #STATUS_TEACH_DYNAMIC_BUSY;

                               IF #teachFunction = #TEACH_FUNCTION_1 AND #statMyPermitTeach1 THEN
                                   // Start Teach
                                   #statRwRecordIOLData[0] := #TICMD_TEACH_SP_START;
                               ELSIF #teachFunction = #TEACH_FUNCTION_2 AND #statMyPermitTeach2 AND #statTeachStarted THEN
                                   // Stop Teach
                                   #statRwRecordIOLData[0] := #TICMD_TEACH_SP_STOP;
                               END_IF;

                               #statFBSubState := #FB_SUB_STATE_DYNAMIC_WRITE_COMMAND;
                           END_IF;

                           // Send Stop Teach Command if time is up
                           IF #statTeachStarted AND #teachTimer <> T#0ms AND #instTimer.Q = TRUE THEN
                               // Stop Teach
                               #statRwRecordIOLData[0] := #TICMD_TEACH_SP_STOP;
                               #statFBSubState := #FB_SUB_STATE_DYNAMIC_WRITE_COMMAND;
                           END_IF;

                           // Update status information
                           IF #statFBSubState = #FB_SUB_STATE_DYNAMIC_UPDATE_STATUS THEN
                               #instDevice(execute := TRUE,
                                           readWrite := #MODE_READ,
                                           index := #INDEX_TI_RESULT,
                                           record := #statRwRecordIOLData);

                               IF #instDevice.done THEN
                                   #instDevice(execute := FALSE,
                                               record := #statRwRecordIOLData);

                                   // Evaluate response from device
                                   IF (#statRwRecordIOLData[0] AND #MASK_TEACH_STATE) = INT_TO_BYTE(#TEACH_STATE_IDLE) OR
                                       (#statRwRecordIOLData[0] AND #MASK_TEACH_STATE) = INT_TO_BYTE(#TEACH_STATE_SUCCESS)
                                   THEN // Idle and success are handled as error because wait for command is expected here
                                       #statStatus := #ERR_TEACH_DEVICE;
                                   ELSIF (#statRwRecordIOLData[0] AND #MASK_TEACH_STATE) = INT_TO_BYTE(#TEACH_STATE_WAIT_FOR_COMMAND) THEN
                                       #statStatus := #STATUS_TEACH_DYNAMIC_WAITING;
                                       #statFBSubState := 0;
                                       #statTeachStarted := TRUE;
                                       #statMyPermitTeach1 := FALSE;
                                       #statMyPermitTeach2 := TRUE;
                                       #statMyPermitAbort := TRUE;
                                   ELSIF (#statRwRecordIOLData[0] AND #MASK_TEACH_STATE) = INT_TO_BYTE(#TEACH_STATE_BUSY) THEN
                                       #statStatus := #STATUS_TEACH_DYNAMIC_BUSY;
                                   ELSIF (#statRwRecordIOLData[0] AND #MASK_TEACH_STATE) = INT_TO_BYTE(#TEACH_STATE_ERROR) THEN
                                       #statStatus := #ERR_TEACH_DEVICE;
                                   ELSE
                                       #statStatus := #ERR_TEACH_DEVICE;
                                   END_IF;
                               END_IF;
                           END_IF;

                           IF #statFBSubState = #FB_SUB_STATE_DYNAMIC_WRITE_COMMAND THEN
                               #instDevice(execute := TRUE,
                                           readWrite := #MODE_WRITE,
                                           index := #INDEX_SYS_CMD,
                                           writeLen := 1,
                                           record := #statRwRecordIOLData);

                               IF #instDevice.done THEN
                                   #instDevice(execute := FALSE,
                                               record := #statRwRecordIOLData);

                                   IF #statRwRecordIOLData[0] = #TICMD_TEACH_SP_START THEN
                                       #statFBSubState := #FB_SUB_STATE_DYNAMIC_UPDATE_STATUS;

                                       // Start Teach Timer
                                       IF #teachTimer <> T#0ms THEN
                                           #instTimer(PT := #teachTimer,
                                                      IN := TRUE);
                                       END_IF;

                                   ELSIF #statRwRecordIOLData[0] = #TICMD_TEACH_SP_STOP THEN
                                       #statFBState := #FB_STATE_CHECK_RESULT;
                                       #statStatus := #STATUS_TEACH_APPLYING; // Busy, Teach process, apply action
                                   END_IF;

                                   #statMyPermitAbort := TRUE;
                               END_IF;
                           END_IF;
                       END_IF;
                   END_REGION dynamic teach-in

                   REGION check result
                       IF #statFBState = #FB_STATE_CHECK_RESULT THEN
                           #statMyPermitTeach1 := FALSE;
                           #statMyPermitTeach2 := FALSE;
                           #statMyPermitApply := FALSE;
                           #statMyPermitAbort := FALSE;

                           // Read Teach-in state
                           #instDevice(execute := TRUE,
                                       readWrite := #MODE_READ,
                                       index := #INDEX_TI_RESULT,
                                       record := #statRwRecordIOLData);

                           IF #instDevice.done THEN
                               #instDevice(execute := FALSE,
                                           record := #statRwRecordIOLData);

                               IF (#statRwRecordIOLData[0] AND #MASK_TEACH_STATE) = INT_TO_BYTE(#TEACH_STATE_BUSY) THEN
                                   ; // Keep trying until teach state of device is not busy
                               ELSIF (#statRwRecordIOLData[0] AND #MASK_TEACH_STATE) = INT_TO_BYTE(#TEACH_STATE_SUCCESS) THEN
                                   #statMyPermitTeach1 := FALSE;
                                   #statMyPermitTeach2 := FALSE;
                                   #statMyPermitApply := FALSE;
                                   #statMyPermitAbort := FALSE;

                                   #statFBState := #FB_STATE_READ_ALL; // Go to read all
                                   #statIndexRead := #INDEX_SSC_PARAM;
                                   #statLenRead := 2;
                               ELSIF (#statRwRecordIOLData[0] AND #MASK_TEACH_STATE) = INT_TO_BYTE(#TEACH_STATE_WAIT_FOR_COMMAND) THEN
                                   #statStatus := #STATUS_TEACH_WAITING_APPLY;
                               ELSIF (#statRwRecordIOLData[0] AND #MASK_TEACH_STATE) = INT_TO_BYTE(#TEACH_STATE_ERROR) THEN
                                   #statStatus := #ERR_TEACH_DEVICE;
                               END_IF;
                           END_IF;
                       END_IF;
                   END_REGION check result

                   REGION abort
                       // Check for Abort Teach and not permitted Functions
                       IF #teachRequest AND NOT #statTeachRequestOld THEN
                           IF #teachFunction = #TEACH_FUNCTION_1 AND NOT #statMyPermitTeach1
                               OR #teachFunction = #TEACH_FUNCTION_2 AND NOT #statMyPermitTeach2
                               OR #teachFunction = #TEACH_FUNCTION_APPLY AND NOT #statMyPermitApply
                               OR #teachFunction = #TEACH_FUNCTION_ABORT AND NOT #statMyPermitAbort THEN
                               #statStatus := #ERR_TEACH_NOT_ALLOWED;
                           ELSIF #teachFunction = #TEACH_FUNCTION_ABORT AND #statMyPermitAbort THEN
                               #statFBState := #FB_STATE_ABORT_TEACH;
                           END_IF;
                       END_IF;

                       IF #statFBState = #FB_STATE_ABORT_TEACH THEN
                           #statStatus := #STATUS_TEACH_ABORTING;

                           // Abort Teach-in sequence
                           #statRwRecordIOLData[0] := #TICMD_TEACH_CANCEL;
                           #instDevice(execute := TRUE,
                                       readWrite := #MODE_WRITE,
                                       index := #INDEX_SYS_CMD,
                                       writeLen := 1,
                                       record := #statRwRecordIOLData);

                           IF #instDevice.done THEN
                               #instDevice(execute := FALSE,
                                           record := #statRwRecordIOLData);

                               #statStatus := #STATUS_EXECUTION_FINISHED;
                           END_IF;
                       END_IF;
                   END_REGION abort

                   // Error Handling
                   IF #instDevice.error THEN
                       #statStatus := #ERR_DEVICE_FB;
                       #statSubfunctionStatus := #instDevice.status;
                       #statFBErrorState := #statFBSubState;
                   END_IF;
               END_REGION teach

           #FB_STATE_READ_ALL..#FB_STATE_BACKUP:
               REGION param exchange
                   // State to read and write Setpoint and Logic

                   REGION read all
                       IF #statFBState = #FB_STATE_READ_ALL THEN // Read "Logic" and "Setpoint"
                           #statStatus := #STATUS_BUSY_READING; // Busy reading data

                           #instDevice(execute := TRUE,
                                       readWrite := #MODE_READ,
                                       index := #statIndexRead,
                                       record := #statRwRecordIOLData);

                           IF #instDevice.done THEN
                               #instDevice(execute := FALSE,
                                           record := #statRwRecordIOLData);

                               IF #statIndexRead >= #INDEX_SSC_CONFIG THEN
                                   #logicOut := BYTE_TO_BOOL(#statRwRecordIOLData[0] AND 2#00000001);

                                   IF #backupEnable AND #function = #FUNC_TEACH THEN
                                       #statFBState := #FB_STATE_BACKUP;
                                   ELSE
                                       #statStatus := #STATUS_EXECUTION_FINISHED;
                                   END_IF;

                               ELSE
                                   #tempSetpointOut1.%B0 := #statRwRecordIOLData[1];
                                   #tempSetpointOut1.%B1 := #statRwRecordIOLData[0];
                                   #setpointOut1 := WORD_TO_INT(#tempSetpointOut1);

                                   #tempSetpointOut2.%B0 := #statRwRecordIOLData[1];
                                   #tempSetpointOut2.%B1 := #statRwRecordIOLData[0];
                                   #setpointOut2 := WORD_TO_INT(#tempSetpointOut2);

                                   // Read "Logic" after reading "Setpoint"
                                   #statIndexRead += 1;
                                   #statLenRead := 1;
                               END_IF;
                           END_IF;
                       END_IF;
                   END_REGION read all

                   REGION write config
                       IF #statFBState = #FB_STATE_WRITE_CONF THEN
                           #statStatus := #STATUS_BUSY_WRITING; // Busy writing data
                           #statRwRecordIOLData[0] := BOOL_TO_BYTE(#logicIn);

                           #instDevice(execute := true,
                                       readWrite := #MODE_WRITE,
                                       index := #INDEX_SSC_CONFIG,
                                       writeLen := 1,
                                       record := #statRwRecordIOLData);

                           IF #instDevice.done THEN
                               //Write input to output if writing was successful
                               #logicOut := #logicIn;

                               IF #backupEnable THEN
                                   #statFBState := #FB_STATE_BACKUP;
                                   #instDevice(execute := FALSE,
                                               record := #statRwRecordIOLData);
                               ELSE
                                   #statStatus := #STATUS_EXECUTION_FINISHED;
                               END_IF;
                           END_IF;
                       END_IF;
                   END_REGION write config

                   REGION write param
                       IF #statFBState = #FB_STATE_WRITE_PARAM THEN
                           #statStatus := #STATUS_BUSY_WRITING;

                           #tempSetpointIn1 := INT_TO_WORD(#setpointIn1);
                           #statRwRecordIOLData[1] := #tempSetpointIn1.%B0;
                           #statRwRecordIOLData[0] := #tempSetpointIn1.%B1;

                           #tempSetpointIn2 := INT_TO_WORD(#setpointIn2);
                           #statRwRecordIOLData[1] := #tempSetpointIn2.%B0;
                           #statRwRecordIOLData[0] := #tempSetpointIn2.%B1;

                           #instDevice(execute := TRUE,
                                       readWrite := #MODE_WRITE,
                                       index := #INDEX_SSC_PARAM,
                                       writeLen := 2,
                                       record := #statRwRecordIOLData);

                           IF #instDevice.done THEN
                               //Write input to output if writing was successful
                               #setpointOut1 := #setpointIn1;
                               #setpointOut2 := #setpointIn2;
                               IF #backupEnable THEN
                                   #statFBState := #FB_STATE_BACKUP;
                                   #instDevice(execute := FALSE,
                                               record := #statRwRecordIOLData);
                               ELSE
                                   #statStatus := #STATUS_EXECUTION_FINISHED;
                               END_IF;
                           END_IF;
                       END_IF;
                   END_REGION write param

                   REGION param download store
                       IF #statFBState = #FB_STATE_BACKUP THEN
                           #statStatus := #STATUS_BUSY_BACKUP; // Busy backup
                           #statRwRecordIOLData[0] := 16#05;

                           #instDevice(execute := TRUE,
                                       readWrite := #MODE_WRITE,
                                       index := #INDEX_SYS_CMD,
                                       writeLen := 1,
                                       record := #statRwRecordIOLData);

                           IF #instDevice.done THEN
                               #statStatus := #STATUS_EXECUTION_FINISHED;
                           END_IF;
                       END_IF;
                   END_REGION param download store

                   // Error handling
                   IF #instDevice.error THEN
                       #statStatus := #ERR_DEVICE_FB;
                       #statSubfunctionStatus := #instDevice.status;
                       #statFBErrorState := #statFBState;
                   END_IF;
               END_REGION param exchange
       END_CASE;
   END_REGION STATE_MACHINE

   REGION OUTPUTS
       // Write outputs
       IF (#statStatus = #STATUS_EXECUTION_FINISHED) AND (#statDone = FALSE) THEN // Execution finished without errors
           REGION execution finished
               #statDone := TRUE;
               #statBusy := FALSE;
               #statError := FALSE;

               #statMyPermitTeach1 := FALSE;
               #statMyPermitTeach2 := FALSE;
               #statMyPermitApply := FALSE;
               #statMyPermitAbort := FALSE;

               // execution aborted --> set state no processing
               #statFBState := #FB_STATE_NO_PROCESSING;
               #statFBState := 0;
               #statFBSubState := 0;
           END_REGION execution finished

       ELSIF (#statStatus.%X15 = TRUE) AND (#statError = FALSE) THEN // Error occurred (#statStatus is 16#8000 to 16#FFFF)
           REGION error occured
               #statDone := FALSE;
               #statBusy := FALSE;
               #statError := TRUE;

               #statMyPermitTeach1 := FALSE;
               #statMyPermitTeach2 := FALSE;
               #statMyPermitApply := FALSE;
               #statMyPermitAbort := FALSE;

               // Write diagnostics
               #diagnostics.status := #statStatus;
               #diagnostics.subfunctionStatus := #statSubfunctionStatus;
               #diagnostics.stateNumber := #statFBErrorState;

               // Reset instance for next job
               #instDevice(execute := FALSE,
                           record := #statRwRecordIOLData);

               // execution aborted --> set state no processing
               #statFBState := #FB_STATE_NO_PROCESSING;
               #statFBState := 0;
               #statFBSubState := 0;
           END_REGION error occured

       ELSIF (#tempExecute = FALSE) AND ((#statDone = TRUE) OR (#statError = TRUE)) THEN // Reset outputs
           REGION execute reset
               #statDone := FALSE;
               #statBusy := FALSE;
               #statError := FALSE;
               #statStatus := #STATUS_NO_CALL;

               // Reset instance for next job
               #instDevice(execute := FALSE,
                           record := #statRwRecordIOLData);

           END_REGION execute reset
       END_IF;

       REGION Write static values to outputs
           #done := #statDone;
           #busy := #statBusy;
           #error := #statError;
           #status := #statStatus;

           // Write internal used variables to outputs
           #permitTeach1 := #statMyPermitTeach1;
           #permitTeach2 := #statMyPermitTeach2;
           #permitApply := #statMyPermitApply;
           #permitAbort := #statMyPermitAbort;

           // Needed to detect rising edge at inputs
           #statTeachRequestOld := #teachRequest;

           ENO := NOT #statError;
       END_REGION Write static values to outputs
   END_REGION OUTPUTS
END_FUNCTION_BLOCK

FUNCTION_BLOCK "LIOLink_MeasuredDataChannel"   // FB9, SCL
TITLE = IOL_MeasurementDataChannel / LIOLink_MeasuringDataChannel
{ S7_Optimized_Access := 'TRUE' }
AUTHOR : SUP_Applications
FAMILY : LIOLink
VERSION : 1.0
// The Measurement Data Channel defines the Process Data structure, functions and representation of measuring sensors. This Function Block provides derived status signals and defines a standardized interface for user application programs. If this FB is migrated to another automation system, than the input measurementValue of type Variant probably has to be replaced by a suitable alternative.
   VAR_INPUT
      profileID : Word;   // 1 = SSP 3.1; 2 = SSP 3.2; 3 = SSP 3.3; 4 = SSP 3.4 / 1 = SSP 3.1; 2 = SSP 3.2; 3 = SSP 3.3; 4 = SSP 3.4; 5 = SSP 4.1.x; 6 = SSP 4.2.x
      substituteValue : DInt;   // This value is applied at the outputs ValueReal and Val-ueDINT if ValueStatus is not equal 0
      qualifier : Bool;   // false = ProcessData are invalid; true = ProcessData are valid
      LogicStartAddress : Int;   // Logical address of the first byte from Process Data input structure
   END_VAR
   VAR_OUTPUT
      valid : Bool;   // If “true” the provided values are valid and may be used for further calculations
      error : Bool;   // If “true” an internal error is occurred and futher information is provided provided by the Function Block via the Status variable
      status : Word := 16#0000;   // Provides internal error codes
      valueStatus : Int;   // Status of process data input: 0 = OK; 1 = PC invalid; 2 = No Data; 3 = Out of range (+); 4 = Out of range (-); 5 = Not defined
      valueReal : Real;   // Process data in real format for evaluation within the PLC
      valueDInt : DInt;   // Process data in double integer format
      scale : Int;   // Process data scale factor
      "SSCn.1" : Bool;   // Switching information channel 1
      "SSCn.2" : Bool;   // Switching information channel 2
   END_VAR
   VAR_TEMP
      iScale : SInt;   // Scale information from process image
      byScale : Byte;   // Scale information from process image
      iMeasurementValue : Int;   // Measurement Value as Integer
      wMeasurementValue : Word;   // Measurement Value as Word
      diMeasurementValue : DInt;   // Measurement Value as Double Integer
      dwMeasurementValue : DWord;   // Measurement Value as Double Word
   END_VAR
   VAR CONSTANT
      LOWER_LIMIT_INT : Int := -32768;   // Value which represents lower limit of 16 bit measurement value
      UPPER_LIMIT_INT : Int := 32767;   // Value which represents upper limit of 16 bit measurement value
      LOWER_LIMIT_DINT : DInt := -2147482880;   // Value which represents lower limit of 32 bit measurement value
      UPPER_LIMIT_DINT : DInt := 2147482880;   // Value which represents upper limit of 32 bit measurement value
      OUT_OF_RANGE_NEG_INT : Int := 16#8008;   // Value which represents that 16 bit measurement value is out of range (-)
      OUT_OF_RANGE_POS_INT : Int := 16#7FF8;   // Value which represents that 16 bit measurement value is out of range (+)
      OUT_OF_RANGE_NEG32 : DInt := 16#80000008;   // Value which represents that 32 bit measurement value is out of range (-)
      OUT_OF_RANGE_POS32 : DInt := 16#7FFFFFF8;   // Value which represents that 32 bit measurement value is out of range (+)
      NO_MEASUREMENT_DATA16 : Int := 16#7FFC;   // Value which represents that IOL_Device cannot provide a 16 bit measurement value
      NO_MEASUREMENT_DATA32 : DInt := 16#7FFFFFFC;   // Value which represents that IOL_Device cannot provide a 32 bit measurement value
      VAL_STAT_OK : Int := 0;   // Value for Status = OK
      VAL_STAT_PD_INVALID : Int := 1;   // Value for Status = Process Data invalid
      VAL_STAT_NO_DATA : Int := 2;   // Value for Status = No Data
      VAL_STAT_OUT_OF_RANGE_POS : Int := 3;   // Value for Status = Measurement Value out of range (-)
      VAL_STAT_OUT_OF_RANGE_NEG : Int := 4;   // Value for Status = Measurement Value out of range (+)
      VAL_STAT_NOT_DEFINED : Int := 5;   // Value for Status = Measurement Value not defined
      ERR_UNDEFINED_PROFILE_ID : DWord := 16#00000001;   // Error code for unvalid ProfileId at input / Status Code if the value at input ProfileId is not defined
      STATUS_READY_TO_START : Word := 16#0000;   // Status: Teach process successfull/ Ready to Start Teach-In process / idle / Status: Order completed, no warning
      STATUS_UNKNOWN_PROFIL_ID : Word := 16#8001;   // Status: An unknown profil ID is used
      PROFILID_SSP1 : Word := 1;   // Profil ID=1, SSP 3.1
      PROFILID_SSP2 : Word := 2;   // Profil ID=2, SSP 3.2
      PROFILID_SSP3 : Word := 3;   // Profil ID=3, SSP 3.3
      PROFILID_SSP4 : Word := 4;   // Profil ID=4, SSP 3.4
      PROFILID_SSP5 : Word := 5;   // Profil ID=4, SSP 3.4
      PROFILID_SSP6 : Word := 6;
   END_VAR
BEGIN
   REGION BLOCK INFO HEADER
     //===============================================================================
     // Siemens / (c)Copyright 2020
     //-------------------------------------------------------------------------------
     // Title:            LIOLink_MeasuredDataChannel
     // Function:         The Measurement Data Channel defines the Process Data         
     //                   structure, functions and representation of measuring sensors.   
     //                   This Function Block provides derived status signals and            
     //                   defines a standardized interface for user application programs. 
     // Library:          LIOLink
     // Author:           SUP Applications
     // Tested with:      CPU 1513-1 PN FW 2.8
     // Engineering:      TIA Portal V16
     // Restrictions:     --
     // Requirements:     --
     //-------------------------------------------------------------------------------
     // Change log table:
     // Version  | Date       | Expert in charge       | Changes applied
     //----------|------------|------------------------|------------------------------
     // 01.00.00 | 06.03.2019 | SUP Applications       | First release
     // 01.00.04 | 22.09.2020 | Online Support         | Enabled block simulation support
     // 02.00.00 | 31.03.2023 | SUP Applications       | Added support of SSP 4.1.x and SSP 4.2.x                      
     //                                                 Replaced input "MeasurementValue" (Variant) by                
     //                                                 "LogicStartAddress" (INT)                                     
     //                                                 Removed input ScaleIn                                         
     //                                                 Added outputs SSCn.1 and SSCn.2
     //===============================================================================
   END_REGION

   REGION Init outputs
       #error := FALSE;
       #status := #STATUS_READY_TO_START;
       #"SSCn.1" := 0;
       #"SSCn.2" := 0;
   END_REGION

   REGION Init temp variables
       #iScale := 0;
       #byScale := 0;
       #iMeasurementValue := 0;
       #wMeasurementValue := 0;
       #diMeasurementValue := 0;
       #dwMeasurementValue := 0;
   END_REGION

   IF #qualifier = FALSE THEN
     #valueDInt := #substituteValue;
     #valueReal := DINT_TO_REAL(#substituteValue);
     #valueStatus := #VAL_STAT_PD_INVALID;
     #valid := FALSE;

   ELSE
     //SSP 3.1 or 3.3 or 4.1.x
       IF (#profileID = #PROFILID_SSP1 OR #profileID = #PROFILID_SSP3 OR #profileID = #PROFILID_SSP5) THEN
           REGION 16-bit measurement value 
               #wMeasurementValue := PEEK_WORD(area := 16#81, dbNumber := 0, byteOffset := #LogicStartAddress);
               #iMeasurementValue := WORD_TO_INT(#wMeasurementValue);
               #byScale := PEEK(area := 16#81, dbNumber := 0, byteOffset := #LogicStartAddress + 2);
               #iScale := BYTE_TO_SINT(#byScale);

               IF #profileID = #PROFILID_SSP5 THEN
                   #"SSCn.1" := PEEK_BOOL(area := 16#81, dbNumber := 0, byteOffset := #LogicStartAddress + 3, bitOffset := 0);
                   #"SSCn.2" := PEEK_BOOL(area := 16#81, dbNumber := 0, byteOffset := #LogicStartAddress + 3, bitOffset := 1);
               END_IF;

               IF #LOWER_LIMIT_INT <= #iMeasurementValue AND #iMeasurementValue <= #UPPER_LIMIT_INT THEN
                   #valueDInt := #iMeasurementValue;
                   #valueReal := INT_TO_REAL(#iMeasurementValue) * (10 ** INT_TO_REAL(#iScale));
                   #valueStatus := #VAL_STAT_OK;
                   #valid := TRUE;

               ELSE
                   IF #iMeasurementValue = #OUT_OF_RANGE_POS_INT THEN
                       #valueStatus := #VAL_STAT_OUT_OF_RANGE_POS;

                   ELSIF #iMeasurementValue = #OUT_OF_RANGE_NEG_INT THEN
                       #valueStatus := #VAL_STAT_OUT_OF_RANGE_NEG;

                   ELSIF #iMeasurementValue = #NO_MEASUREMENT_DATA16 THEN
                       #valueStatus := #VAL_STAT_NO_DATA;

                   ELSE // MeasurementValue does not fit any defined Value
                       #valueStatus := #VAL_STAT_NOT_DEFINED;

                   END_IF;
                   #valueDInt := #substituteValue;
                   #valueReal := DINT_TO_REAL(#substituteValue);
                   #valid := FALSE;
               END_IF;
           END_REGION
       //SSP 3.2 or 3.4 or 4.2.x
   ELSIF (#profileID = #PROFILID_SSP2 OR #profileID = #PROFILID_SSP4 OR #profileID = #PROFILID_SSP6) THEN
       REGION 32-bit measurement value
           #dwMeasurementValue := PEEK_DWORD(area := 16#81, dbNumber := 0, byteOffset := #LogicStartAddress);
           #diMeasurementValue := DWORD_TO_DINT(#dwMeasurementValue);
           #byScale := PEEK(area := 16#81, dbNumber := 0, byteOffset := #LogicStartAddress + 4);
           #iScale := BYTE_TO_SINT(#byScale);

           IF #profileID = #PROFILID_SSP6 THEN
               #"SSCn.1" := PEEK_BOOL(area := 16#81, dbNumber := 0, byteOffset := #LogicStartAddress + 5, bitOffset := 0);
               #"SSCn.2" := PEEK_BOOL(area := 16#81, dbNumber := 0, byteOffset := #LogicStartAddress + 5, bitOffset := 1);
           END_IF;

           IF #LOWER_LIMIT_DINT <= #diMeasurementValue AND #diMeasurementValue <= #UPPER_LIMIT_DINT THEN
               #valueDInt := #diMeasurementValue;
               #valueReal := DINT_TO_REAL(#diMeasurementValue) * (10 ** INT_TO_REAL(#iScale));
               #valueStatus := #VAL_STAT_OK;
               #valid := TRUE;

           ELSE
               IF #diMeasurementValue = #OUT_OF_RANGE_POS32 THEN
                   #valueStatus := #VAL_STAT_OUT_OF_RANGE_POS;

               ELSIF #diMeasurementValue = #OUT_OF_RANGE_NEG32 THEN
                   #valueStatus := #VAL_STAT_OUT_OF_RANGE_NEG;

               ELSIF #diMeasurementValue = #NO_MEASUREMENT_DATA32 THEN
                   #valueStatus := #VAL_STAT_NO_DATA;

               ELSE // MeasurementValue does not fit any defined Value
                   #valueStatus := #VAL_STAT_NOT_DEFINED;
               END_IF;

               #valueDInt := #substituteValue;
               #valueReal := DINT_TO_REAL(#substituteValue);
               #valid := FALSE;
           END_IF;
       END_REGION
     ELSE  // Statement section ELSE
       #valueDInt := #substituteValue;
       #valueReal := DINT_TO_REAL(#substituteValue);
       #valueStatus := #VAL_STAT_OK;
       #valid := FALSE;
       #error := TRUE;
       #status := #STATUS_UNKNOWN_PROFIL_ID;
     END_IF;
   END_IF;

   #scale := #iScale;
END_FUNCTION_BLOCK

// folder: Profile blocks

